(* CODESYS project PersistentVars.gvl.xml

Project tree, tasks and I/O mapping:
  global variables PersistentVars
*)

// PersistentVars
{attribute 'qualified_only'}
VAR_GLOBAL PERSISTENT RETAIN
	// Generated instance path of persistent variable
	PLC_PRG.Alarm.Settings: ST_AlarmSettings;
	// Generated instance path of persistent variable
	PLC_PRG.Alarm.Configuration: ST_AlarmHmiConfiguration;
END_VAR
